// TIA Portal V20 export
// export: Created 2026-10-06T00:00:00
Screen "Conveyor_Settings"  1280x800, Number=3, Template=Base
  ScreenLayer 
    Rectangle "Speed" at 30,100 size 40x40
